Fanuc KAREL source: kt00301.KL

-- PROVISIONAL review KL for V1013-1; original PC SHA256 7d8220d8ebb3db5cfb62dfe440b63fbe94bd9ee0eaf28d05bb26fa83749b8ddb
-- Incomplete behavior may be omitted. Consult companion uncertainty JSON. Do not deploy.
PROGRAM KT00301
%NOLOCKGROUP
VAR
  B1 : BOOLEAN
  B2 : BOOLEAN
  OUT : BOOLEAN
BEGIN
  -- UNRESOLVED_PC offsets 5-12; opcodes 9D,23
  -- UNRESOLVED_PC offsets 17-24; opcodes 9C,23
  -- UNRESOLVED_PC offsets 29-36; opcodes 9D,23
  -- UNRESOLVED_PC offsets 41-48; opcodes 9C,23
  -- UNRESOLVED_PC offsets 53-72; opcodes 21,21,58,23
  -- UNRESOLVED_PC offsets 77-81; opcodes 7F
END KT00301
